Fanuc KAREL source: kt00437.KL

-- PROVISIONAL review KL for V1013-1; original PC SHA256 40648883f964a363df25fca36df8198ee29af265f16d55e8ed149f822c11b21a
-- Incomplete behavior may be omitted. Consult companion uncertainty JSON. Do not deploy.
PROGRAM KT00437
%NOLOCKGROUP
VAR
  I1 : INTEGER
  I2 : INTEGER
  OUT : BOOLEAN
BEGIN
  -- UNRESOLVED_PC offsets 5-16; opcodes 2E,23
  -- UNRESOLVED_PC offsets 21-32; opcodes 2E,23
  -- UNRESOLVED_PC offsets 37-48; opcodes 2E,23
  -- UNRESOLVED_PC offsets 53-64; opcodes 2E,23
  -- UNRESOLVED_PC offsets 69-88; opcodes 21,21,5C,23
  -- UNRESOLVED_PC offsets 93-97; opcodes 7F
END KT00437
